{region 'Documentation'}
(*!
<summary>Checks that selected bits match the expected masked value.</summary>
*)
{endregion}
FUNCTION_BLOCK AssertEqualMask_Byte EXTENDS AssertionBase
VAR_INPUT
    IN : BYTE; //! Actual bitfield.
    Mask : BYTE := 16#FF; //! Selects evaluated bits; defaults to all bits. An empty mask produces Error during evaluation.
    Expected : BYTE; //! Expected value; bits outside Mask are ignored.
END_VAR

SUPER^();

{region 'Documentation'}
(*!
<summary>Rejects an empty mask before comparing selected bits.</summary>
*)
{endregion}
METHOD PROTECTED Assert
VAR
    Message : STRING(GVL_Constants.MessageLength);
    MaskText : STRING(GVL_Constants.AssertionValueLength);
    ExpectedText : STRING(GVL_Constants.AssertionValueLength);
    ActualText : STRING(GVL_Constants.AssertionValueLength);
END_VAR
VAR CONSTANT
    NoMask : BYTE := 16#00;
    HexDigitCount : USINT := 2;
END_VAR
IF NOT EvaluationActive THEN
    RETURN;
END_IF;

IF Result = E_Result.Error THEN
    RETURN;
END_IF;

IF Mask = NoMask THEN
    MaskText := CreateAssertionTextValue_Hex(Value := BYTE_TO_LWORD(Mask),
        DigitCount := HexDigitCount);
    Message := CONCAT('Assertion error: mask must not be empty. Mask = ',
        MaskText);
    Message := CONCAT(Message, '.');
    Error(Message := Message);
    RETURN;
END_IF;

IF Result = E_Result.Failed THEN
    RETURN;
END_IF;

IF (IN AND Mask) <> (Expected AND Mask) THEN
    MaskText := CreateAssertionTextValue_Hex(Value := BYTE_TO_LWORD(Mask),
        DigitCount := HexDigitCount);
    ExpectedText := CreateAssertionTextValue_Hex(Value := BYTE_TO_LWORD(Expected),
        DigitCount := HexDigitCount);
    ActualText := CreateAssertionTextValue_Hex(Value := BYTE_TO_LWORD(IN),
        DigitCount := HexDigitCount);
    Message := CONCAT('Assertion failed: selected bits do not match. Expected = ',
        ExpectedText);
    Message := CONCAT(Message, ', Mask = ');
    Message := CONCAT(Message, MaskText);
    Message := CONCAT(Message, ', Actual = ');
    Message := CONCAT(Message, ActualText);
    Message := CONCAT(Message, '.');
    Fail(Message := Message);
    RETURN;
END_IF;

Pass();
END_METHOD

END_FUNCTION_BLOCK

(* stored: Version 1.1.0.1
   POU AssertEqualMask_Byte: Id {fa3d9517-b19f-462d-8a71-099219dfee79}, SpecialFunc None
   Folder Internal: Id {a48ea389-13a3-4713-9ef5-7e7cb22aaa46}
   Method Assert: Id {74dcf1a5-3e32-4e2a-a267-d3f44cb02c5b} *)
